TYPE "ST_UnitProbeDevice"
VERSION : 0.1
   STRUCT
      Cycles : UDInt;
      ExitCalls : UDInt;
      Changes : UDInt;
      Resets : UDInt;
      Received : Bool;
      Processed : Bool;
   END_STRUCT;

END_TYPE

